TYPE stLightConfig :
STRUCT
	BrightnessRamp : BOOL := FALSE;
	BrightnessRampTime : TIME := T#2S;
END_STRUCT
END_TYPE

(* stored: Version 1.1.0.1
   DUT stLightConfig: Id {52e1058c-f365-49f2-9c9d-7fb722dfb0a0} *)
